Fanuc KAREL source: ka00122.KL

-- PROVISIONAL review KL for V770-1; original PC SHA256 5121194bc6c395452ec271c8408275fff88aa036f6349413134f70c81b521b65
-- Incomplete behavior may be omitted. Consult companion uncertainty JSON. Do not deploy.
PROGRAM KA00122
%NOLOCKGROUP
VAR
  DST : REAL
-- UNRESOLVED_DECL SRC type=002018
BEGIN
  -- UNRESOLVED_PC offsets 5-19; opcodes 2E,22,9D,33,B2
  -- UNRESOLVED_PC offsets 24-40; opcodes 22,9D,33,B1,64,23
  -- UNRESOLVED_PC offsets 45-49; opcodes 7F
END KA00122
